Staubli VAL3: trajectory.dtx

mdesc mNomSpeed
frame fFrame = {fatherId=world[0]}
tool tTool = {fatherId=flange[0]}
mdesc mSim = {blend=off}
frame _fFrame = {fatherId=world[0]}
pointRx pGOTO = {fatherId=world[0]}
num nIndex[100]
